// ============================================================================
// DB_TestBench: 测试台背景数据块 (FB_9001_TestBench_DJ2026011 的实例 DB)
// 说明: 背景 DB 不写变量, 变量来自 FB; 由 OB 调用测试台时使用。
// ============================================================================

DATA_BLOCK "DB_TestBench"
"FB_9001_TestBench_DJ2026011"
BEGIN
END_DATA_BLOCK
